Fanuc KAREL source: KA00051.KL

PROGRAM KA00051
%NOLOCKGROUP
VAR
  SRC: POSITION
  DST: BOOLEAN
BEGIN
  DST = SRC
END KA00051
